Fanuc KAREL source: ka00120.KL

-- PROVISIONAL review KL for V770-1; original PC SHA256 f0edb6afc8a94cdcdc43c4b0d560b9d0c9da7df76b539037a25893a9cca8ccfe
-- Incomplete behavior may be omitted. Consult companion uncertainty JSON. Do not deploy.
PROGRAM KA00120
%NOLOCKGROUP
-- UNRESOLVED_DECL SRC type=00001c
-- UNRESOLVED_DECL DST type=002017
BEGIN
  -- UNRESOLVED_PC offsets 5-15; opcodes 9D,22,A5
  -- UNRESOLVED_PC offsets 20-35; opcodes 21,22,9D,33,B4
  -- UNRESOLVED_PC offsets 40-44; opcodes 7F
END KA00120
